FUNCTION_BLOCK LineModule EXTENDS ModuleGroup
VAR
    _Filler           : I_EquipmentModule;
    _Transfer         : I_EquipmentModule;
    _State            : E_LineState;
    _IsStartRequested : BOOL;
    _IsStopping       : BOOL;
    _IsConfigured     : BOOL;
END_VAR
(*
    LineModule

    The machine module. Fills a bottle, moves it out, and repeats until
    stopped. Commands its two stations in BeforeChildren(), before they
    run in the same scan.

    Start() starts the line. Stop() lets the bottle in progress finish.
    A fault anywhere in the tree stops commanding and shows Faulted; once
    the tree no longer reports a fault, the line is Stopped and waits for
    Start(). Reset(), inherited, resets the whole tree.
*)

METHOD FB_init : BOOL
VAR_INPUT
    bInitRetains : BOOL;
    bInCopyCode  : BOOL;
    Name         : STRING(32);                  // for EquipmentGroup
    Filler       : I_EquipmentModule;
    Transfer     : I_EquipmentModule;
END_VAR
_Filler := Filler;
_Transfer := Transfer;
_IsConfigured := Filler <> 0 AND Transfer <> 0;
END_METHOD

METHOD PUBLIC Start
_IsStartRequested := TRUE;
_IsStopping := FALSE;                           // a start cancels a stop that hasn't been taken yet
END_METHOD

METHOD PUBLIC Stop
IF _State <> E_LineState.Stopped THEN
    _IsStopping := TRUE;                        // taken when the bottle is out
END_IF
END_METHOD

METHOD PROTECTED BeforeChildren
IF NOT _IsConfigured THEN
    _State := E_LineState.Faulted;
    RETURN;
END_IF

// A fault anywhere in the tree: command nothing
IF HasFault THEN
    _State := E_LineState.Faulted;
    _IsStopping := FALSE;
    _IsStartRequested := FALSE;
    RETURN;
END_IF

CASE _State OF
    E_LineState.Stopped:
        IF _IsStartRequested THEN
            _Filler.StartCycle();
            _State := E_LineState.Filling;
        END_IF

    E_LineState.Filling:
        IF _Filler.IsCycleDone THEN
            _Transfer.StartCycle();
            _State := E_LineState.Transferring;
        END_IF

    E_LineState.Transferring:
        IF _Transfer.IsCycleDone THEN
            IF _IsStopping THEN
                _IsStopping := FALSE;
                _State := E_LineState.Stopped;
            ELSE
                _Filler.StartCycle();           // the next bottle
                _State := E_LineState.Filling;
            END_IF
        END_IF

    E_LineState.Faulted:
        _State := E_LineState.Stopped;          // no fault any more; wait for Start
END_CASE

_IsStartRequested := FALSE;
END_METHOD

PROPERTY PUBLIC State : E_LineState
GET
State := _State;
END_GET
END_PROPERTY

PROPERTY PUBLIC IsStopping : BOOL
GET
IsStopping := _IsStopping;
END_GET
END_PROPERTY

END_FUNCTION_BLOCK

(* stored: Version 1.1.0.1, ProductVersion 3.1.4026.0
   POU LineModule: Id {af7f9873-6eef-4792-929d-8b412e3c19b2}, SpecialFunc None
   Method FB_init: Id {a3e47bab-b4fc-4fdc-ac0f-e91f9b4bf2d0}
   Method Start: Id {b51082b5-7bf0-4ac5-985a-ceb9b9a57dfb}
   Method Stop: Id {cb6d3e2e-d34a-456d-b08f-3760254f7239}
   Method BeforeChildren: Id {7e3d8405-7c71-40d1-a594-92fa05f9416f}
   Property State: Id {e74d5d94-e787-4e84-a09f-db1dfef1e31e}
   Get Get: Id {80350595-bef7-4fe2-8874-a5730eaac171}
   Property IsStopping: Id {9766d7e4-70ee-4d9d-9910-50212f3d24a6}
   Get Get: Id {dac68dd1-70a6-447a-9797-d7392f6a4a26} *)
